Staubli VAL3: setPage.pgx

public program setPage(num x_nType)
begin
  switch x_nType
    case 0,1

      nPage=roundUp(io:nMaxdigital/16)

    break
    case 2,3
      nPage=roundUp(io:nMaxAnalog/16)
      if nPageIndex>nPage-1
        nPageIndex=0
      endIf
    break
  endSwitch
  sPageNum=toString("",nPage)
  sShowPageIndex=toString("",nPageIndex+1)
end
